Staubli VAL3: refreshCheckBox.pgx

public program refreshCheckBox(utImage& x_utImage[])
  local num l_nI
  local num l_nJ
begin
    if size(x_utImage) != 1
      for l_nI= 0 to size(x_utImage)-1
        if x_utImage[l_nI].Events.bClick==true
          x_utImage[l_nI].Events.bClick=false
          l_nJ=l_nI
          for l_nI=0 to size(x_utImage)-1
            if l_nI==l_nJ
              x_utImage[l_nI].Common.sSourceImage=x_utImage[l_nI].Data.sSourceImg1
              x_utImage[l_nI].Data.bStatus=true
            else
              x_utImage[l_nI].Common.sSourceImage=x_utImage[l_nI].Data.sSourceImg2
              x_utImage[l_nI].Data.bStatus=false
            endIf
          endFor
        endIf
      endFor
    else
      if x_utImage[l_nI].Events.bClick==true
        x_utImage[l_nI].Events.bClick=false
        if x_utImage[l_nI].Data.bStatus==false
          x_utImage[l_nI].Common.sSourceImage=x_utImage[l_nI].Data.sSourceImg1
          x_utImage[l_nI].Data.bStatus=true
        else
          x_utImage[l_nI].Common.sSourceImage=x_utImage[l_nI].Data.sSourceImg2
          x_utImage[l_nI].Data.bStatus=false
        endIf
      endIf
    endIf
end
